PROGRAM prg_Call_OpMode
VAR
	fbModeMain:FB_ModeSelect;
	
	rt_HMI_Resume: R_TRIG;
	rt_ActError: R_TRIG;
	
	eModeZone: E_ModeZone;

END_VAR

fbModeMain(sModuleDescription:='Mode Select - Main',
	bInterlockBypass:=TRUE, //bIntZoneBypass[1]
	bLockedFB:=TRUE, //bIntZoneLocked[1]
	bPistonCheck:=FALSE,	
	bLockRequest=>,	//bReq_LockZone[1]
	eModeZone:=E_ModeZone.eMain,
	stMode:=stModeMain,
	stOperation:=stOpMain, 
	bStateSafe_mode:=bStateSafe);
	
FOR eModeZone:=	E_ModeZone.eMain TO E_ModeZone.eLast DO
	fbMode[eModeZone](sModuleDescription:='Mode Select - ',
		bInterlockBypass:=TRUE, //bIntZoneBypass[eModeZone]
		bLockedFB:=TRUE, //bIntZoneLocked[eModeZone]
		bPistonCheck:=FALSE,	
		bLockRequest=>,	//bReq_LockZone[eModeZone]
		eModeZone:=eModeZone,
		stMode:=stMode[eModeZone],
		stOperation:=stOper[eModeZone],
		bStateSafe_mode:=m_Get_StateSafe_by_ModeZone(eMoZone:=eModeZone));	
END_FOR
	
PauseAll:=stOpMain.iActOperation=E_OperationButtons.ePauseAll;	
PauseAllDelayed:=stOpMain.bPauseOnDelayed;	

stOpNonPause.iActOperation:=E_OperationButtons.ePlayAll;
	
rt_HMI_Resume(CLK:=ResumeAll);
IF rt_HMI_Resume.Q THEN;
	stOpMain.bSetPlay:=TRUE;
	prg_Messages.act_ResumeSFC();	
	FOR eModeZone:=	E_ModeZone.eMain TO E_ModeZone.eLast DO;
		stOper[eModeZone].bSetPlay:=TRUE;
	END_FOR
END_IF
ResumeAll:=FALSE;

rt_ActError(CLK:=iActErrors<>0);
IF iActErrors<>0 THEN;
	stOpMain.bSetPause:=TRUE;
END_IF

prg_LightTower(
	bBuzzerBypass:=bBuzzerMute , 
	qLedGreen=> , //q_EL16[2].ch11
	qLedYellow=> , //q_EL16[2].ch10
	qLedRed=> , //q_EL16[2].ch9
	qBuzzer=> );//q_EL16[2].ch12
	
	
act_Call_LightTowers();

ACTION act_Call_LightTowers:
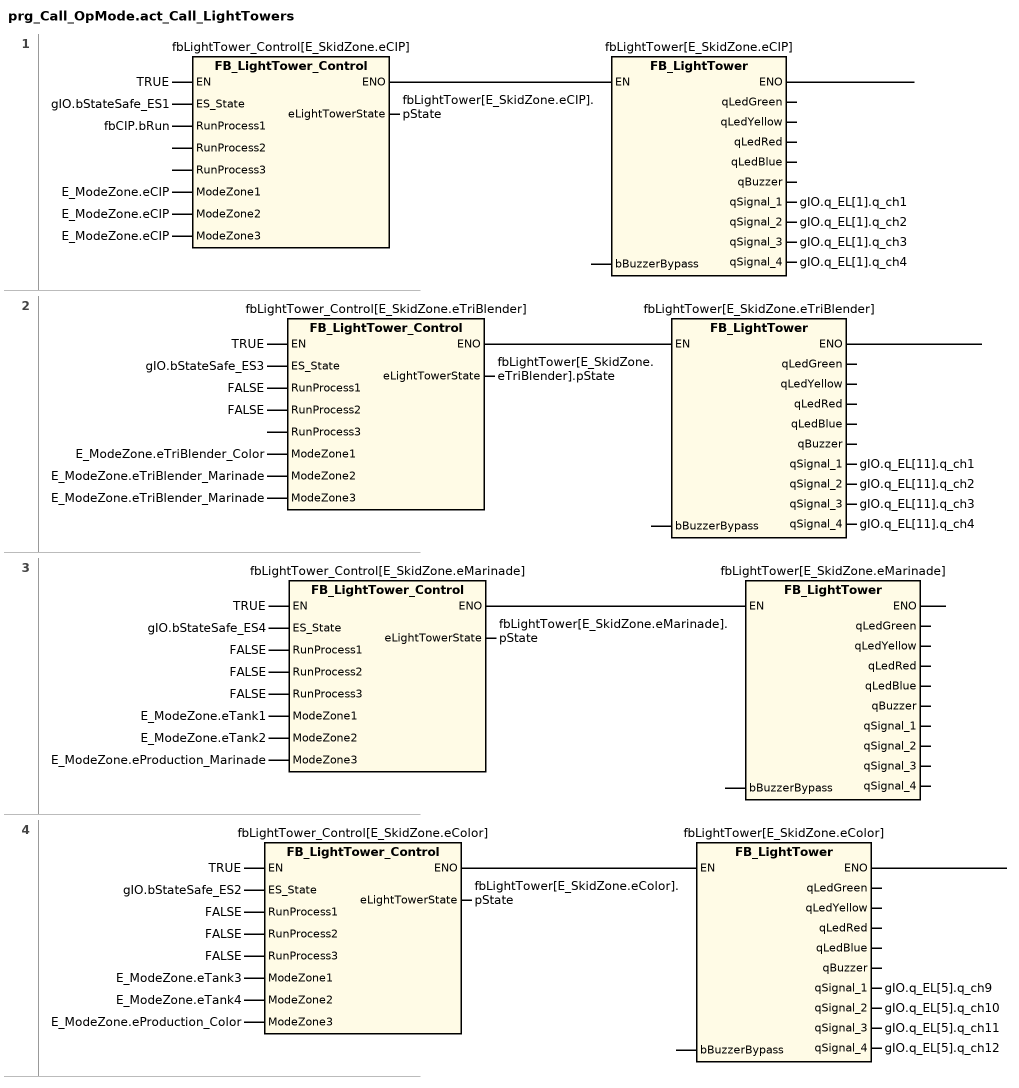
// NETWORK 1
fbLightTower_Control[E_SkidZone.eCIP](
    ES_State := gIO.bStateSafe_ES1,
    RunProcess1 := fbCIP.bRun,
    ModeZone1 := E_ModeZone.eCIP,
    ModeZone2 := E_ModeZone.eCIP,
    ModeZone3 := E_ModeZone.eCIP,
    eLightTowerState => fbLightTower[E_SkidZone.eCIP].pState); // FB_LightTower_Control
fbLightTower[E_SkidZone.eCIP](
    qSignal_1 => gIO.q_EL[1].q_ch1,
    qSignal_2 => gIO.q_EL[1].q_ch2,
    qSignal_3 => gIO.q_EL[1].q_ch3,
    qSignal_4 => gIO.q_EL[1].q_ch4); // FB_LightTower

// NETWORK 2
fbLightTower_Control[E_SkidZone.eTriBlender](
    ES_State := gIO.bStateSafe_ES3,
    RunProcess1 := FALSE,
    RunProcess2 := FALSE,
    ModeZone1 := E_ModeZone.eTriBlender_Color,
    ModeZone2 := E_ModeZone.eTriBlender_Marinade,
    ModeZone3 := E_ModeZone.eTriBlender_Marinade,
    eLightTowerState => fbLightTower[E_SkidZone.eTriBlender].pState); // FB_LightTower_Control
fbLightTower[E_SkidZone.eTriBlender](
    qSignal_1 => gIO.q_EL[11].q_ch1,
    qSignal_2 => gIO.q_EL[11].q_ch2,
    qSignal_3 => gIO.q_EL[11].q_ch3,
    qSignal_4 => gIO.q_EL[11].q_ch4); // FB_LightTower

// NETWORK 3
fbLightTower_Control[E_SkidZone.eMarinade](
    ES_State := gIO.bStateSafe_ES4,
    RunProcess1 := FALSE,
    RunProcess2 := FALSE,
    RunProcess3 := FALSE,
    ModeZone1 := E_ModeZone.eTank1,
    ModeZone2 := E_ModeZone.eTank2,
    ModeZone3 := E_ModeZone.eProduction_Marinade,
    eLightTowerState => fbLightTower[E_SkidZone.eMarinade].pState); // FB_LightTower_Control
fbLightTower[E_SkidZone.eMarinade](); // FB_LightTower

// NETWORK 4
fbLightTower_Control[E_SkidZone.eColor](
    ES_State := gIO.bStateSafe_ES2,
    RunProcess1 := FALSE,
    RunProcess2 := FALSE,
    RunProcess3 := FALSE,
    ModeZone1 := E_ModeZone.eTank3,
    ModeZone2 := E_ModeZone.eTank4,
    ModeZone3 := E_ModeZone.eProduction_Color,
    eLightTowerState => fbLightTower[E_SkidZone.eColor].pState); // FB_LightTower_Control
fbLightTower[E_SkidZone.eColor](
    qSignal_1 => gIO.q_EL[5].q_ch9,
    qSignal_2 => gIO.q_EL[5].q_ch10,
    qSignal_3 => gIO.q_EL[5].q_ch11,
    qSignal_4 => gIO.q_EL[5].q_ch12); // FB_LightTower
END_ACTION

METHOD INTERNAL m_Get_StateSafe_by_ModeZone : BOOL
VAR_INPUT
	eMoZone: E_ModeZone;
END_VAR
CASE eMoZone OF
	E_ModeZone.eCIP:;
		m_Get_StateSafe_by_ModeZone:=bStateSafe_ES1;

	E_ModeZone.eTank3,
	E_ModeZone.eTank4,
	E_ModeZone.eProduction_Color:;
		m_Get_StateSafe_by_ModeZone:=bStateSafe_ES2;		

	E_ModeZone.eTriBlender_Color,
	E_ModeZone.eTriBlender_Marinade:;
		m_Get_StateSafe_by_ModeZone:=bStateSafe_ES3;
		
	E_ModeZone.eTank1,
	E_ModeZone.eTank2,
	E_ModeZone.eProduction_Marinade:;
		m_Get_StateSafe_by_ModeZone:=bStateSafe_ES4;
		
ELSE;
		m_Get_StateSafe_by_ModeZone:=FALSE;
		
END_CASE
(*
bStateSafe_ES1:=arSafe[1].stSafetyIn.ES1_State;
bStateSafe_ES2:=arSafe[1].stSafetyIn.ES2_State;
bStateSafe_ES3:=arSafe[1].stSafetyIn.ES3_State;
bStateSafe_ES4:=arSafe[1].stSafetyIn.ES4_State;
*)
END_METHOD

END_PROGRAM

(* stored: Version 1.1.0.1, ProductVersion 3.1.4024.15
   POU prg_Call_OpMode: Id {37ea252d-f7d6-4416-870e-8e42ec6784ac}, SpecialFunc None
   Action act_Call_LightTowers: Id {7558a2c9-c3f1-4401-ba46-b92b27544782}
   Method m_Get_StateSafe_by_ModeZone: Id {fdafcf64-1d55-4ecf-a98a-8debd67a4d40} *)
